FUNCTION_BLOCK FB_Device
VAR_INPUT
	{attribute 'OPC.UA.DA' := '1'}
	{attribute 'OPC.UA.DA.StructuredType' := '1'}
	ctrl : ST_DeviceControl;
	parentCtrl : ST_ParentChildControl;
END_VAR
VAR_OUTPUT
	{attribute 'instance-path'}
	{attribute 'no-init'}
	instancePath		: T_MaxString;
END_VAR
VAR
	bInit : BOOL := TRUE;

	parentConfigured : BOOL;
	
	{attribute 'hide'} 
	opActivity 		 : BOOL; 
	{attribute 'OPC.UA.DA' := '1'}
	{attribute 'OPC.UA.DA.Access' := '1'} // read only
	{attribute 'OPC.UA.DA.StructuredType' := '1'}
	manualOvrdeTimer : TON;
	{attribute 'hide'} 
	lastMode		 : E_SystemMode := E_SystemMode.Manual;
	{attribute 'hide'} 
	rtModeChange	 : BOOL; 
	{attribute 'hide'} 
	rtBypass		 : R_TRIG;
	{attribute 'hide'} 
	ftBypass	  	 : F_TRIG;
	{attribute 'hide'} 
	rtSim			 : R_TRIG;
	{attribute 'hide'} 
	ftSim			 : F_TRIG;
	
	//------ Configuration ------//
	// Hidden because the cfg variable in the extending 
	// FB will act as a passthrough to these.
	{attribute 'hide'} 
	opTimeout : TIME;
	{attribute 'hide'} 
	opTimeoutEnable : BOOL;
	
	//---------- Status ---------//
	// Hidden because the sts variable in the extending 
	// FB will pass these back out to the user.
	{attribute 'hide'} 
	mode : E_SystemMode := E_SystemMode.Manual;
END_VAR

IF bInit THEN
	Init();
	bInit := FALSE;
END_IF

parentConfigured := parentCtrl.instancePath <> '';

manualOvrdeTimer(IN := ctrl.manualOvrde AND NOT opActivity, PT := opTimeout);
IF manualOvrdeTimer.Q AND opTimeoutEnable THEN
	ctrl.manualOvrde := FALSE;
END_IF

// Determine device mode
CASE mode OF
	E_SystemMode.Idle:
		// Device is switched off locally. Enter/leave this state based on the status of a
		// physical switch co-located with the device. Not implemented yet.
	E_SystemMode.Auto:
		IF ctrl.manualOvrde	OR (parentConfigured AND parentCtrl.mode <> E_SystemMode.Auto) THEN
			mode := E_SystemMode.Manual;
		END_IF
	E_SystemMode.Manual:									
		IF NOT ctrl.manualOvrde AND (NOT parentConfigured OR parentCtrl.mode = E_SystemMode.Auto) THEN
			mode := E_SystemMode.Auto;
		END_IF
	ELSE
		mode := E_SystemMode.Idle;
END_CASE
rtModeChange := mode <> lastMode;
lastMode := mode;

// Triggers
rtBypass(CLK := ctrl.bypass);
ftBypass(CLK := ctrl.bypass);
rtSim(CLK := ctrl.sim);
ftSim(CLK := ctrl.sim);

METHOD PUBLIC DisableBypass
ctrl.bypass := FALSE;
END_METHOD

METHOD PUBLIC DisableManualOverride
ctrl.manualOvrde := FALSE;
END_METHOD

METHOD PUBLIC DisableSimulation
ctrl.sim := FALSE;
END_METHOD

METHOD PUBLIC EnableBypass
ctrl.bypass := TRUE;
END_METHOD

METHOD PUBLIC EnableManualOverride
ctrl.manualOvrde := TRUE;
END_METHOD

METHOD PUBLIC EnableSimulation
ctrl.sim := TRUE;
END_METHOD

METHOD PROTECTED Init : BOOL
// Insert code here that must be completed before function block runs.
// Set output conditionally based on this code
Init := TRUE;
END_METHOD

METHOD PUBLIC Reset
ctrl.reset := TRUE;
END_METHOD

END_FUNCTION_BLOCK

(* stored: Version 1.1.0.1, ProductVersion 3.1.4024.12
   POU FB_Device: Id {3365eada-ff13-41a7-bfcc-aef33150f2ed}, SpecialFunc None
   Folder Control: Id {8079e94b-57e8-4684-98c3-75435637ba16}
   Method DisableBypass: Id {83d963cb-2f77-466b-89e6-ced59503c491}
   Method DisableManualOverride: Id {2dd37739-9e89-4d33-b18c-1335f68b673e}
   Method DisableSimulation: Id {5920d782-0e41-4241-af6c-3fd227461b68}
   Method EnableBypass: Id {2da2c4de-ec2e-4df7-b307-e4d0020cc2bb}
   Method EnableManualOverride: Id {8eb69e79-c413-4ede-8059-31e4f2dcf6a9}
   Method EnableSimulation: Id {6edd7fae-1a72-4baf-add9-141f62e72d55}
   Method Init: Id {c8498a5a-bddd-4405-bf14-0201ed8de335}
   Method Reset: Id {b7f79351-370a-47c8-8ba9-cb76c2204640} *)
